// TIA Portal V19 export
VAR_GLOBAL   // PLC tag table "R1_IN"
   "ByteIN :0 R1" AT %IB90 : Byte;   // System Bits 1
   "ByteIN :1 R1" AT %IB91 : Byte;   // System Bits 2
   "ByteIN :2 R1" AT %IB92 : Byte;   // Signals
   "ByteIN :3 R1" AT %IB93 : Byte;   // Signals
   "ByteIN :4 R1" AT %IB94 : Byte;   // CMD
   "ByteIN :5 R1" AT %IB95 : Byte;
   "ByteIN :6 R1" AT %IB96 : Byte;
   "ByteIN :7 R1" AT %IB97 : Byte;
   "ByteIN :8 R1" AT %IB98 : Byte;
   "ByteIN :9 R1" AT %IB99 : Byte;
   "ByteIN :10 R1" AT %IB100 : Byte;
   "ByteIN :11 R1" AT %IB101 : Byte;
   "ByteIN :12 R1" AT %IB102 : Byte;
   "ByteIN :13 R1" AT %IB103 : Byte;
   "ByteIN :14 R1" AT %IB104 : Byte;
   "ByteIN :15 R1" AT %IB105 : Byte;
   "ByteIN :16 R1" AT %IB106 : Byte;
   "ByteIN :17 R1" AT %IB107 : Byte;
   "ByteIN :18 R1" AT %IB108 : Byte;
   "ByteIN :19 R1" AT %IB109 : Byte;
   "ByteIN :20 R1" AT %IB110 : Byte;
   "ByteIN :21 R1" AT %IB111 : Byte;
   "ByteIN :22 R1" AT %IB112 : Byte;
   "ByteIN :23 R1" AT %IB113 : Byte;
   "ByteIN :24 R1" AT %IB114 : Byte;
   "ByteIN :25 R1" AT %IB115 : Byte;
   "ByteIN :26 R1" AT %IB116 : Byte;
   "ByteIN :27 R1" AT %IB117 : Byte;
   "ByteIN :28 R1" AT %IB118 : Byte;
   "ByteIN :29 R1" AT %IB119 : Byte;
   "ByteIN :30 R1" AT %IB120 : Byte;
   "ByteIN :31 R1" AT %IB121 : Byte;
   "ByteIN :32 R1" AT %IB122 : Byte;
   "ByteIN :33 R1" AT %IB123 : Byte;
   "ByteIN :34 R1" AT %IB124 : Byte;
   "ByteIN :35 R1" AT %IB125 : Byte;
   "ByteIN :36 R1" AT %IB126 : Byte;
   "ByteIN :37 R1" AT %IB127 : Byte;
   "ByteIN :38 R1" AT %IB128 : Byte;
   "ByteIN :39 R1" AT %IB129 : Byte;
   "ByteIN :40 R1" AT %IB130 : Byte;
   "ByteIN :41 R1" AT %IB131 : Byte;
   "ByteIN :42 R1" AT %IB132 : Byte;
   "ByteIN :43 R1" AT %IB133 : Byte;
   "ByteIN :44 R1" AT %IB134 : Byte;
   "ByteIN :45 R1" AT %IB135 : Byte;
   "ByteIN :46 R1" AT %IB136 : Byte;
   "ByteIN :47 R1" AT %IB137 : Byte;
   "ByteIN :48 R1" AT %IB138 : Byte;
   "ByteIN :49 R1" AT %IB139 : Byte;
   "ByteIN :50 R1" AT %IB140 : Byte;
   "ByteIN :51 R1" AT %IB141 : Byte;
   "ByteIN :52 R1" AT %IB142 : Byte;
   "ByteIN :53 R1" AT %IB143 : Byte;
   "ByteIN :54 R1" AT %IB144 : Byte;
   "ByteIN :55 R1" AT %IB145 : Byte;
   "ByteIN :56 R1" AT %IB146 : Byte;
   "ByteIN :57 R1" AT %IB147 : Byte;
   "ByteIN :58 R1" AT %IB148 : Byte;
   "ByteIN :59 R1" AT %IB149 : Byte;
   "ByteIN :60 R1" AT %IB150 : Byte;
   "ByteIN :61 R1" AT %IB151 : Byte;
   "ByteIN :62 R1" AT %IB152 : Byte;
   "ByteIN :63 R1" AT %IB153 : Byte;
END_VAR
